Staubli VAL3: kill.pgx

program kill()
begin
  //kill all task
  taskKill("safeCheck")
  taskKill("Reset")
  taskKill("Start")
  taskKill("Stop")
  taskKill("cycleCtrl")
  taskKill("plc")
  taskKill("lifebit")
  taskKill("actCtrl")
  taskKill("appMain")
  taskKill("HMI")

  //
  rs:bQuitApp=false
  stopMove()
  resetMotion()
  disablePower()
end
